(* IEC 61131-3 sources: PortalRobot/Portal_robot/Device/application/ST/ST_GRIPPER, 7 files *)

(* ---- E_GRIPPER_STATE.st ---- *)
{attribute 'qualified_only'}
{attribute 'strict'}
TYPE E_GRIPPER_STATE :
(
	IDLE,
    EXECUTE,
    DONE,
    ERROR
);
END_TYPE

(* ---- ST_GRIPPER_COMMAND.st ---- *)
TYPE ST_GRIPPER_COMMAND :
STRUCT
	xExecute : BOOL; // Команда запуска действия
	xReset   : BOOL; // Команда сброса ошибки
	eAction  : E_ROBOT_ACTION; // Требуемое действие захвата
	// Дискретный контракт исполнительных механизмов. Каждый BOOL задаёт
	// состояние своего механизма: 0 — закрыть/к заготовке, 1 — открыть/к детали.
	xGripper1Open   : BOOL; // Захват 1: 0 закрыть, 1 открыть
	xGripper2Open   : BOOL; // Захват 2: 0 закрыть, 1 открыть
	xRotateToDetail : BOOL; // Поворот: 0 к заготовке, 1 к детали
END_STRUCT
END_TYPE

(* ---- ST_GRIPPER_DIAG.st ---- *)
TYPE ST_GRIPPER_DIAG :
STRUCT
	eState        : E_GRIPPER_STATE; // Текущее состояние автомата
	eActiveAction : E_ROBOT_ACTION; // Выполняемое действие захвата
	stWarning     : ST_WARNING_EVENT; // Последнее предупреждение захвата
END_STRUCT
END_TYPE

(* ---- ST_GRIPPER_ERROR.st ---- *)
TYPE ST_GRIPPER_ERROR :
STRUCT
	GRIPPER_1_ERROR : BOOL; // Ошибка первого захвата
	GRIPPER_2_ERROR : BOOL; // Ошибка второго захвата
	ROTATION_ERROR  : BOOL; // Ошибка механизма поворота
	ACTION_ERROR    : BOOL; // Получено недопустимое действие
	GLOBAL_ERROR    : BOOL; // Глобальная ошибка симуляции захвата
END_STRUCT
END_TYPE

(* ---- ST_GRIPPER_ERRORS.st ---- *)
TYPE ST_GRIPPER_ERRORS :
STRUCT
	dwErrorActive : DWORD; // Битовая маска активных ошибок
	dwErrorLast   : DWORD; // Битовая маска последних ошибок
	dwAlarmActive : DWORD; // Собственные аварии захвата для общего журнала
	stErrorActive : ST_GRIPPER_ERROR; // Расшифровка активных ошибок
	stErrorLast   : ST_GRIPPER_ERROR; // Расшифровка последних ошибок
END_STRUCT
END_TYPE

(* ---- ST_GRIPPER_FAULT_REQUEST.st ---- *)
TYPE ST_GRIPPER_FAULT_REQUEST :
STRUCT
	xEnabled        : BOOL; // Глобальное разрешение диагностической инъекции
	xGripper1Fault  : BOOL; // Неисправность первого захвата
	xGripper2Fault  : BOOL; // Неисправность второго захвата
	xRotationFault  : BOOL; // Неисправность механизма поворота
	xGlobalFault    : BOOL; // Общая неисправность захвата
END_STRUCT
END_TYPE

(* ---- ST_GRIPPER_STATUS.st ---- *)
TYPE ST_GRIPPER_STATUS  :
STRUCT
	xBusy            : BOOL; // Выполняется действие захвата
	xDone            : BOOL; // Действие завершено
	xError           : BOOL; // Захват находится в ошибке
	xGripper1Open    : BOOL; // Первый захват открыт
	xGripper1Closed  : BOOL; // Первый захват закрыт
	xGripper2Open    : BOOL; // Второй захват открыт
	xGripper2Closed  : BOOL; // Второй захват закрыт
	xRotatedToBlank  : BOOL; // Захват повёрнут к заготовке
	xRotatedToDetail : BOOL; // Захват повёрнут к детали
END_STRUCT
END_TYPE
